(* IEC 61131-3 sources: matiec/tests/initialization, 38 files *)

(* ---- bad_array_nested_too_many_outer.st ---- *)
(* Test of initial values for structured/array data types. *)

TYPE
  arr_dint : ARRAY [1..2] OF DINT;
  arr_arr_dint : ARRAY [1..2] OF arr_dint;
END_TYPE

PROGRAM program0
  VAR
    count : DINT;
    v : arr_arr_dint := [[1, 2], [3, 4], [5, 6]];
  END_VAR

  count := count + 1;
END_PROGRAM

CONFIGURATION config
  RESOURCE resource1 ON PLC
    TASK main_task(INTERVAL := T#1000ms, PRIORITY := 0);
    PROGRAM instance0 WITH main_task : program0;
  END_RESOURCE
END_CONFIGURATION

(* ---- bad_array_scalar_for_struct_element.st ---- *)
(* Test of initial values for structured/array data types. *)

TYPE
  inner : STRUCT
    a : DINT;
    b : DINT;
    c : STRING;
  END_STRUCT;
  arr_inner : ARRAY [1..2] OF inner;
END_TYPE

PROGRAM program0
  VAR
    count : DINT;
    v : arr_inner := [5, 6];
  END_VAR

  count := count + 1;
END_PROGRAM

CONFIGURATION config
  RESOURCE resource1 ON PLC
    TASK main_task(INTERVAL := T#1000ms, PRIORITY := 0);
    PROGRAM instance0 WITH main_task : program0;
  END_RESOURCE
END_CONFIGURATION

(* ---- bad_array_string_for_scalar_element.st ---- *)
(* Test of initial values for structured/array data types. *)

TYPE
  arr_dint : ARRAY [1..2] OF DINT;
END_TYPE

PROGRAM program0
  VAR
    count : DINT;
    v : arr_dint := ['x', 'y'];
  END_VAR

  count := count + 1;
END_PROGRAM

CONFIGURATION config
  RESOURCE resource1 ON PLC
    TASK main_task(INTERVAL := T#1000ms, PRIORITY := 0);
    PROGRAM instance0 WITH main_task : program0;
  END_RESOURCE
END_CONFIGURATION

(* ---- bad_array_struct_for_scalar_element.st ---- *)
(* Test of initial values for structured/array data types. *)

TYPE
  inner : STRUCT
    a : DINT;
    b : DINT;
    c : STRING;
  END_STRUCT;
  arr_inner : ARRAY [1..2] OF inner;
  arr_dint : ARRAY [1..2] OF DINT;
END_TYPE

PROGRAM program0
  VAR
    count : DINT;
    v : arr_dint := [(a := 1, b := 2, c := 'a'), (a := 3, b := 4, c := 'b')];
  END_VAR

  count := count + 1;
END_PROGRAM

CONFIGURATION config
  RESOURCE resource1 ON PLC
    TASK main_task(INTERVAL := T#1000ms, PRIORITY := 0);
    PROGRAM instance0 WITH main_task : program0;
  END_RESOURCE
END_CONFIGURATION

(* ---- bad_array_too_many_in_struct.st ---- *)
(* Test of initial values for structured/array data types. *)

TYPE
  inner : STRUCT
    a : DINT;
    b : DINT;
    c : STRING;
  END_STRUCT;
  arr_inner : ARRAY [1..2] OF inner;
  rec : STRUCT
    kkk : DINT;
    many : arr_inner;
  END_STRUCT;
END_TYPE

PROGRAM program0
  VAR
    count : DINT;
    v : rec := (kkk := 9, many := [(a := 1, b := 2, c := 'a'), (a := 3, b := 4, c := 'b'), (a := 5, b := 6, c := 'e')]);
  END_VAR

  count := count + 1;
END_PROGRAM

CONFIGURATION config
  RESOURCE resource1 ON PLC
    TASK main_task(INTERVAL := T#1000ms, PRIORITY := 0);
    PROGRAM instance0 WITH main_task : program0;
  END_RESOURCE
END_CONFIGURATION

(* ---- bad_array_too_many_multidim.st ---- *)
(* Test of initial values for structured/array data types. *)

TYPE
  arr_dint : ARRAY [1..2, 1..3] OF DINT;
END_TYPE

PROGRAM program0
  VAR
    count : DINT;
    v : arr_dint := [1, 2, 3, 4, 5, 6, 7];
  END_VAR

  count := count + 1;
END_PROGRAM

CONFIGURATION config
  RESOURCE resource1 ON PLC
    TASK main_task(INTERVAL := T#1000ms, PRIORITY := 0);
    PROGRAM instance0 WITH main_task : program0;
  END_RESOURCE
END_CONFIGURATION

(* ---- bad_array_too_many_nested.st ---- *)
(* Test of initial values for structured/array data types. *)

TYPE
  arr_dint : ARRAY [1..2] OF DINT;
  arr_arr_dint : ARRAY [1..2] OF arr_dint;
END_TYPE

PROGRAM program0
  VAR
    count : DINT;
    v : arr_arr_dint := [[1, 2], [3, 4, 5]];
  END_VAR

  count := count + 1;
END_PROGRAM

CONFIGURATION config
  RESOURCE resource1 ON PLC
    TASK main_task(INTERVAL := T#1000ms, PRIORITY := 0);
    PROGRAM instance0 WITH main_task : program0;
  END_RESOURCE
END_CONFIGURATION

(* ---- bad_array_too_many_of_struct.st ---- *)
(* Test of initial values for structured/array data types. *)

TYPE
  inner : STRUCT
    a : DINT;
    b : DINT;
    c : STRING;
  END_STRUCT;
  arr_inner : ARRAY [1..2] OF inner;
END_TYPE

PROGRAM program0
  VAR
    count : DINT;
    v : arr_inner := [(a := 1, b := 2, c := 'a'), (a := 3, b := 4, c := 'b'), (a := 5, b := 6, c := 'e')];
  END_VAR

  count := count + 1;
END_PROGRAM

CONFIGURATION config
  RESOURCE resource1 ON PLC
    TASK main_task(INTERVAL := T#1000ms, PRIORITY := 0);
    PROGRAM instance0 WITH main_task : program0;
  END_RESOURCE
END_CONFIGURATION

(* ---- bad_array_too_many_repeated.st ---- *)
(* Test of initial values for structured/array data types. *)

TYPE
  arr_dint : ARRAY [1..2] OF DINT;
END_TYPE

PROGRAM program0
  VAR
    count : DINT;
    v : arr_dint := [4(7)];
  END_VAR

  count := count + 1;
END_PROGRAM

CONFIGURATION config
  RESOURCE resource1 ON PLC
    TASK main_task(INTERVAL := T#1000ms, PRIORITY := 0);
    PROGRAM instance0 WITH main_task : program0;
  END_RESOURCE
END_CONFIGURATION

(* ---- bad_array_too_many_values.st ---- *)
(* Test of initial values for structured/array data types. *)

TYPE
  arr_dint : ARRAY [1..2] OF DINT;
END_TYPE

PROGRAM program0
  VAR
    count : DINT;
    v : arr_dint := [1, 2, 3];
  END_VAR

  count := count + 1;
END_PROGRAM

CONFIGURATION config
  RESOURCE resource1 ON PLC
    TASK main_task(INTERVAL := T#1000ms, PRIORITY := 0);
    PROGRAM instance0 WITH main_task : program0;
  END_RESOURCE
END_CONFIGURATION

(* ---- bad_array_unknown_struct_element.st ---- *)
(* Test of initial values for structured/array data types. *)

TYPE
  inner : STRUCT
    a : DINT;
    b : DINT;
    c : STRING;
  END_STRUCT;
  arr_inner : ARRAY [1..2] OF inner;
END_TYPE

PROGRAM program0
  VAR
    count : DINT;
    v : arr_inner := [(a := 1, zz := 2, c := 'a'), (a := 3, b := 4, c := 'b')];
  END_VAR

  count := count + 1;
END_PROGRAM

CONFIGURATION config
  RESOURCE resource1 ON PLC
    TASK main_task(INTERVAL := T#1000ms, PRIORITY := 0);
    PROGRAM instance0 WITH main_task : program0;
  END_RESOURCE
END_CONFIGURATION

(* ---- bad_struct_array_for_scalar_element.st ---- *)
(* Test of initial values for structured/array data types. *)

TYPE
  arr_dint : ARRAY [1..2] OF DINT;
  rec : STRUCT
    kkk : DINT;
  END_STRUCT;
END_TYPE

PROGRAM program0
  VAR
    count : DINT;
    v : rec := (kkk := [1, 2]);
  END_VAR

  count := count + 1;
END_PROGRAM

CONFIGURATION config
  RESOURCE resource1 ON PLC
    TASK main_task(INTERVAL := T#1000ms, PRIORITY := 0);
    PROGRAM instance0 WITH main_task : program0;
  END_RESOURCE
END_CONFIGURATION

(* ---- bad_struct_scalar_for_struct_element.st ---- *)
(* Test of initial values for structured/array data types. *)

TYPE
  inner : STRUCT
    a : DINT;
    b : DINT;
    c : STRING;
  END_STRUCT;
  rec : STRUCT
    kkk : DINT;
    complex : inner;
  END_STRUCT;
END_TYPE

PROGRAM program0
  VAR
    count : DINT;
    v : rec := (kkk := 1, complex := 5);
  END_VAR

  count := count + 1;
END_PROGRAM

CONFIGURATION config
  RESOURCE resource1 ON PLC
    TASK main_task(INTERVAL := T#1000ms, PRIORITY := 0);
    PROGRAM instance0 WITH main_task : program0;
  END_RESOURCE
END_CONFIGURATION

(* ---- bad_struct_unknown_element.st ---- *)
(* Test of initial values for structured/array data types. *)

TYPE
  inner : STRUCT
    a : DINT;
    b : DINT;
    c : STRING;
  END_STRUCT;
END_TYPE

PROGRAM program0
  VAR
    count : DINT;
    v : inner := (a := 1, zz := 2, c := 'a');
  END_VAR

  count := count + 1;
END_PROGRAM

CONFIGURATION config
  RESOURCE resource1 ON PLC
    TASK main_task(INTERVAL := T#1000ms, PRIORITY := 0);
    PROGRAM instance0 WITH main_task : program0;
  END_RESOURCE
END_CONFIGURATION

(* ---- ok_array_enum.st ---- *)
(* Test of initial values for structured/array data types. *)

TYPE
  colour : (RED, GREEN, BLUE);
  arr_colour : ARRAY [1..2] OF colour;
END_TYPE

PROGRAM program0
  VAR
    count : DINT;
    v : arr_colour := [RED, BLUE];
  END_VAR

  count := count + 1;
END_PROGRAM

CONFIGURATION config
  RESOURCE resource1 ON PLC
    TASK main_task(INTERVAL := T#1000ms, PRIORITY := 0);
    PROGRAM instance0 WITH main_task : program0;
  END_RESOURCE
END_CONFIGURATION

(* ---- ok_array_enum_in_typedecl.st ---- *)
(* Test of initial values for structured/array data types. *)

TYPE
  colour : (RED, GREEN, BLUE);
  arr_colour : ARRAY [1..2] OF colour := [RED, BLUE];
END_TYPE

PROGRAM program0
  VAR
    count : DINT;
    v : arr_colour;
  END_VAR

  count := count + 1;
END_PROGRAM

CONFIGURATION config
  RESOURCE resource1 ON PLC
    TASK main_task(INTERVAL := T#1000ms, PRIORITY := 0);
    PROGRAM instance0 WITH main_task : program0;
  END_RESOURCE
END_CONFIGURATION

(* ---- ok_array_fewer_values.st ---- *)
(* Test of initial values for structured/array data types. *)

TYPE
  arr_dint : ARRAY [1..3] OF DINT;
END_TYPE

PROGRAM program0
  VAR
    count : DINT;
    v : arr_dint := [5, 6];
  END_VAR

  count := count + 1;
END_PROGRAM

CONFIGURATION config
  RESOURCE resource1 ON PLC
    TASK main_task(INTERVAL := T#1000ms, PRIORITY := 0);
    PROGRAM instance0 WITH main_task : program0;
  END_RESOURCE
END_CONFIGURATION

(* ---- ok_array_inline_in_struct.st ---- *)
(* Test of initial values for structured/array data types. *)

TYPE
  rec : STRUCT
    kkk : DINT;
    many : ARRAY [1..2] OF DINT;
  END_STRUCT;
END_TYPE

PROGRAM program0
  VAR
    count : DINT;
    v : rec := (kkk := 9, many := [5, 6]);
  END_VAR

  count := count + 1;
END_PROGRAM

CONFIGURATION config
  RESOURCE resource1 ON PLC
    TASK main_task(INTERVAL := T#1000ms, PRIORITY := 0);
    PROGRAM instance0 WITH main_task : program0;
  END_RESOURCE
END_CONFIGURATION

(* ---- ok_array_multidim.st ---- *)
(* Test of initial values for structured/array data types. *)

TYPE
  arr_dint : ARRAY [1..2, 1..3] OF DINT;
END_TYPE

PROGRAM program0
  VAR
    count : DINT;
    v : arr_dint := [1, 2, 3, 4, 5, 6];
  END_VAR

  count := count + 1;
END_PROGRAM

CONFIGURATION config
  RESOURCE resource1 ON PLC
    TASK main_task(INTERVAL := T#1000ms, PRIORITY := 0);
    PROGRAM instance0 WITH main_task : program0;
  END_RESOURCE
END_CONFIGURATION

(* ---- ok_array_nested.st ---- *)
(* Test of initial values for structured/array data types. *)

TYPE
  arr_dint : ARRAY [1..2] OF DINT;
  arr_arr_dint : ARRAY [1..2] OF arr_dint;
END_TYPE

PROGRAM program0
  VAR
    count : DINT;
    v : arr_arr_dint := [[1, 2], [3, 4]];
  END_VAR

  count := count + 1;
END_PROGRAM

CONFIGURATION config
  RESOURCE resource1 ON PLC
    TASK main_task(INTERVAL := T#1000ms, PRIORITY := 0);
    PROGRAM instance0 WITH main_task : program0;
  END_RESOURCE
END_CONFIGURATION

(* ---- ok_array_nested_in_struct.st ---- *)
(* Test of initial values for structured/array data types. *)

TYPE
  arr_dint : ARRAY [1..2] OF DINT;
  arr_arr_dint : ARRAY [1..3] OF arr_dint;
  rec : STRUCT
    kkk : DINT;
    many : arr_arr_dint;
  END_STRUCT;
END_TYPE

PROGRAM program0
  VAR
    count : DINT;
    v : rec := (kkk := 9, many := [[1, 2], [3, 4], [5, 6]]);
  END_VAR

  count := count + 1;
END_PROGRAM

CONFIGURATION config
  RESOURCE resource1 ON PLC
    TASK main_task(INTERVAL := T#1000ms, PRIORITY := 0);
    PROGRAM instance0 WITH main_task : program0;
  END_RESOURCE
END_CONFIGURATION

(* ---- ok_array_nested_in_typedecl.st ---- *)
(* Test of initial values for structured/array data types. *)

TYPE
  arr_dint : ARRAY [1..2] OF DINT;
  arr_arr_dint : ARRAY [1..2] OF arr_dint := [[1, 2], [3, 4]];
END_TYPE

PROGRAM program0
  VAR
    count : DINT;
    v : arr_arr_dint;
  END_VAR

  count := count + 1;
END_PROGRAM

CONFIGURATION config
  RESOURCE resource1 ON PLC
    TASK main_task(INTERVAL := T#1000ms, PRIORITY := 0);
    PROGRAM instance0 WITH main_task : program0;
  END_RESOURCE
END_CONFIGURATION

(* ---- ok_array_nested_inner_partial.st ---- *)
(* Test of initial values for structured/array data types. *)

TYPE
  arr_dint : ARRAY [1..2] OF DINT;
  arr_arr_dint : ARRAY [1..3] OF arr_dint;
END_TYPE

PROGRAM program0
  VAR
    count : DINT;
    v : arr_arr_dint := [[1], [3, 4], [5, 6]];
  END_VAR

  count := count + 1;
END_PROGRAM

CONFIGURATION config
  RESOURCE resource1 ON PLC
    TASK main_task(INTERVAL := T#1000ms, PRIORITY := 0);
    PROGRAM instance0 WITH main_task : program0;
  END_RESOURCE
END_CONFIGURATION

(* ---- ok_array_nested_multidim.st ---- *)
(* Test of initial values for structured/array data types. *)

TYPE
  arr_2d : ARRAY [1..2, 1..3] OF DINT;
  arr_of_2d : ARRAY [1..2] OF arr_2d;
END_TYPE

PROGRAM program0
  VAR
    count : DINT;
    v : arr_of_2d := [[1, 2, 3, 4, 5, 6], [7, 8, 9, 10, 11, 12]];
  END_VAR

  count := count + 1;
END_PROGRAM

CONFIGURATION config
  RESOURCE resource1 ON PLC
    TASK main_task(INTERVAL := T#1000ms, PRIORITY := 0);
    PROGRAM instance0 WITH main_task : program0;
  END_RESOURCE
END_CONFIGURATION

(* ---- ok_array_nested_no_init.st ---- *)
(* Test of initial values for structured/array data types. *)

TYPE
  arr_dint : ARRAY [1..2] OF DINT;
  arr_arr_dint : ARRAY [1..3] OF arr_dint;
END_TYPE

PROGRAM program0
  VAR
    count : DINT;
    v : arr_arr_dint;
  END_VAR

  count := count + 1;
END_PROGRAM

CONFIGURATION config
  RESOURCE resource1 ON PLC
    TASK main_task(INTERVAL := T#1000ms, PRIORITY := 0);
    PROGRAM instance0 WITH main_task : program0;
  END_RESOURCE
END_CONFIGURATION

(* ---- ok_array_nested_of_struct.st ---- *)
(* Test of initial values for structured/array data types. *)

TYPE
  inner : STRUCT
    a : DINT;
    b : DINT;
  END_STRUCT;
  arr_inner : ARRAY [1..2] OF inner;
  arr_arr_inner : ARRAY [1..2] OF arr_inner;
END_TYPE

PROGRAM program0
  VAR
    count : DINT;
    v : arr_arr_inner := [[(a := 1, b := 2), (a := 3, b := 4)], [(a := 5, b := 6), (a := 7, b := 8)]];
  END_VAR

  count := count + 1;
END_PROGRAM

CONFIGURATION config
  RESOURCE resource1 ON PLC
    TASK main_task(INTERVAL := T#1000ms, PRIORITY := 0);
    PROGRAM instance0 WITH main_task : program0;
  END_RESOURCE
END_CONFIGURATION

(* ---- ok_array_nested_partial.st ---- *)
(* Test of initial values for structured/array data types. *)

TYPE
  arr_dint : ARRAY [1..2] OF DINT;
  arr_arr_dint : ARRAY [1..3] OF arr_dint;
END_TYPE

PROGRAM program0
  VAR
    count : DINT;
    v : arr_arr_dint := [[1, 2], [3, 4]];
  END_VAR

  count := count + 1;
END_PROGRAM

CONFIGURATION config
  RESOURCE resource1 ON PLC
    TASK main_task(INTERVAL := T#1000ms, PRIORITY := 0);
    PROGRAM instance0 WITH main_task : program0;
  END_RESOURCE
END_CONFIGURATION

(* ---- ok_array_nested_repeated.st ---- *)
(* Test of initial values for structured/array data types. *)

TYPE
  arr_dint : ARRAY [1..2] OF DINT;
  arr_arr_dint : ARRAY [1..3] OF arr_dint;
END_TYPE

PROGRAM program0
  VAR
    count : DINT;
    v : arr_arr_dint := [3([1, 2])];
  END_VAR

  count := count + 1;
END_PROGRAM

CONFIGURATION config
  RESOURCE resource1 ON PLC
    TASK main_task(INTERVAL := T#1000ms, PRIORITY := 0);
    PROGRAM instance0 WITH main_task : program0;
  END_RESOURCE
END_CONFIGURATION

(* ---- ok_array_of_struct.st ---- *)
(* Test of initial values for structured/array data types. *)

TYPE
  inner : STRUCT
    a : DINT;
    b : DINT;
    c : STRING;
  END_STRUCT;
  arr_inner : ARRAY [1..2] OF inner;
END_TYPE

PROGRAM program0
  VAR
    count : DINT;
    v : arr_inner := [(a := 1, b := 2, c := 'a'), (a := 3, b := 4, c := 'b')];
  END_VAR

  count := count + 1;
END_PROGRAM

CONFIGURATION config
  RESOURCE resource1 ON PLC
    TASK main_task(INTERVAL := T#1000ms, PRIORITY := 0);
    PROGRAM instance0 WITH main_task : program0;
  END_RESOURCE
END_CONFIGURATION

(* ---- ok_array_of_struct_in_struct.st ---- *)
(* Test of initial values for structured/array data types. *)

TYPE
  inner : STRUCT
    a : DINT;
    b : DINT;
    c : STRING;
  END_STRUCT;
  arr_inner : ARRAY [1..2] OF inner;
  rec : STRUCT
    kkk : DINT;
    many : arr_inner;
  END_STRUCT;
END_TYPE

PROGRAM program0
  VAR
    count : DINT;
    v : rec := (kkk := 9, many := [(a := 1, b := 2, c := 'a'), (a := 3, b := 4, c := 'b')]);
  END_VAR

  count := count + 1;
END_PROGRAM

CONFIGURATION config
  RESOURCE resource1 ON PLC
    TASK main_task(INTERVAL := T#1000ms, PRIORITY := 0);
    PROGRAM instance0 WITH main_task : program0;
  END_RESOURCE
END_CONFIGURATION

(* ---- ok_array_of_struct_repeated.st ---- *)
(* Test of initial values for structured/array data types. *)

TYPE
  inner : STRUCT
    a : DINT;
    b : DINT;
    c : STRING;
  END_STRUCT;
  arr_inner : ARRAY [1..2] OF inner;
END_TYPE

PROGRAM program0
  VAR
    count : DINT;
    v : arr_inner := [2((a := 1, b := 2, c := 'a'))];
  END_VAR

  count := count + 1;
END_PROGRAM

CONFIGURATION config
  RESOURCE resource1 ON PLC
    TASK main_task(INTERVAL := T#1000ms, PRIORITY := 0);
    PROGRAM instance0 WITH main_task : program0;
  END_RESOURCE
END_CONFIGURATION

(* ---- ok_array_repeated_value.st ---- *)
(* Test of initial values for structured/array data types. *)

TYPE
  arr_dint : ARRAY [1..4] OF DINT;
END_TYPE

PROGRAM program0
  VAR
    count : DINT;
    v : arr_dint := [2(5), 2(7)];
  END_VAR

  count := count + 1;
END_PROGRAM

CONFIGURATION config
  RESOURCE resource1 ON PLC
    TASK main_task(INTERVAL := T#1000ms, PRIORITY := 0);
    PROGRAM instance0 WITH main_task : program0;
  END_RESOURCE
END_CONFIGURATION

(* ---- ok_array_scalar.st ---- *)
(* Test of initial values for structured/array data types. *)

TYPE
  arr_dint : ARRAY [1..2] OF DINT;
END_TYPE

PROGRAM program0
  VAR
    count : DINT;
    v : arr_dint := [5, 6];
  END_VAR

  count := count + 1;
END_PROGRAM

CONFIGURATION config
  RESOURCE resource1 ON PLC
    TASK main_task(INTERVAL := T#1000ms, PRIORITY := 0);
    PROGRAM instance0 WITH main_task : program0;
  END_RESOURCE
END_CONFIGURATION

(* ---- ok_array_scalar_in_struct.st ---- *)
(* Test of initial values for structured/array data types. *)

TYPE
  arr_dint : ARRAY [1..2] OF DINT;
  rec : STRUCT
    kkk : DINT;
    many : arr_dint;
  END_STRUCT;
END_TYPE

PROGRAM program0
  VAR
    count : DINT;
    v : rec := (kkk := 9, many := [5, 6]);
  END_VAR

  count := count + 1;
END_PROGRAM

CONFIGURATION config
  RESOURCE resource1 ON PLC
    TASK main_task(INTERVAL := T#1000ms, PRIORITY := 0);
    PROGRAM instance0 WITH main_task : program0;
  END_RESOURCE
END_CONFIGURATION

(* ---- ok_array_scalar_in_typedecl.st ---- *)
(* Test of initial values for structured/array data types. *)

TYPE
  arr_dint : ARRAY [1..2] OF DINT := [5, 6];
END_TYPE

PROGRAM program0
  VAR
    count : DINT;
    v : arr_dint;
  END_VAR

  count := count + 1;
END_PROGRAM

CONFIGURATION config
  RESOURCE resource1 ON PLC
    TASK main_task(INTERVAL := T#1000ms, PRIORITY := 0);
    PROGRAM instance0 WITH main_task : program0;
  END_RESOURCE
END_CONFIGURATION

(* ---- ok_struct_element_order.st ---- *)
(* Test of initial values for structured/array data types. *)

TYPE
  inner : STRUCT
    a : DINT;
    b : DINT;
    c : STRING;
  END_STRUCT;
  rec : STRUCT
    kkk : DINT;
    xxx : DINT;
    complex : inner;
  END_STRUCT;
END_TYPE

PROGRAM program0
  VAR
    count : DINT;
    v : rec := (kkk := 1, xxx := 2, complex := (a := 3, b := 4, c := 'a'));
  END_VAR

  count := count + 1;
END_PROGRAM

CONFIGURATION config
  RESOURCE resource1 ON PLC
    TASK main_task(INTERVAL := T#1000ms, PRIORITY := 0);
    PROGRAM instance0 WITH main_task : program0;
  END_RESOURCE
END_CONFIGURATION

(* ---- ok_struct_enum.st ---- *)
(* Test of initial values for structured/array data types. *)

TYPE
  colour : (RED, GREEN, BLUE);
  rec : STRUCT
    kkk : DINT;
    col : colour;
  END_STRUCT;
END_TYPE

PROGRAM program0
  VAR
    count : DINT;
    v : rec := (kkk := 1, col := BLUE);
  END_VAR

  count := count + 1;
END_PROGRAM

CONFIGURATION config
  RESOURCE resource1 ON PLC
    TASK main_task(INTERVAL := T#1000ms, PRIORITY := 0);
    PROGRAM instance0 WITH main_task : program0;
  END_RESOURCE
END_CONFIGURATION

(* ---- ok_struct_nested.st ---- *)
(* Test of initial values for structured/array data types. *)

TYPE
  inner : STRUCT
    a : DINT;
    b : DINT;
    c : STRING;
  END_STRUCT;
  rec : STRUCT
    aa : DINT;
    bb : inner;
  END_STRUCT;
END_TYPE

PROGRAM program0
  VAR
    count : DINT;
    v : rec := (aa := 1, bb := (a := 2, b := 3, c := 'a'));
  END_VAR

  count := count + 1;
END_PROGRAM

CONFIGURATION config
  RESOURCE resource1 ON PLC
    TASK main_task(INTERVAL := T#1000ms, PRIORITY := 0);
    PROGRAM instance0 WITH main_task : program0;
  END_RESOURCE
END_CONFIGURATION
